{region 'Documentation'}
(*!
<summary>Check that IN is strictly later than Minimum.</summary>
*)
{endregion}
FUNCTION_BLOCK AssertLaterThan_Time EXTENDS AssertionBase
VAR_INPUT
    IN : TIME; //! Actual value checked or observed by this Assertion.
    Minimum : TIME; //! Exclusive lower bound; the actual value or count must be greater.
END_VAR

SUPER^();

{region 'Documentation'}
(*!
<summary>Evaluate the typed duration relation and report higher-priority errors first.</summary>
*)
{endregion}
METHOD PROTECTED Assert
VAR
    Message : STRING(GVL_Constants.MessageLength);
    MinimumText : STRING(GVL_Constants.AssertionValueLength);
    ActualText : STRING(GVL_Constants.AssertionValueLength);
END_VAR
IF NOT EvaluationActive THEN
    RETURN;
END_IF;

IF Result = E_Result.Error THEN
    RETURN;
END_IF;

IF Result = E_Result.Failed THEN
    RETURN;
END_IF;

IF IN <= Minimum THEN
    MinimumText := TIME_TO_STRING(Minimum);
    ActualText := TIME_TO_STRING(IN);
    Message := CONCAT('Assertion failed: value is not later than limit. Minimum = ',
        MinimumText);
    Message := CONCAT(Message, ', Actual = ');
    Message := CONCAT(Message, ActualText);
    Message := CONCAT(Message, '.');
    Fail(Message := Message);
    RETURN;
END_IF;

Pass();
END_METHOD

END_FUNCTION_BLOCK

(* stored: Version 1.1.0.1
   POU AssertLaterThan_Time: Id {9ff3d36c-af1e-41ef-b888-d1db9372648d}, SpecialFunc None
   Folder Internal: Id {66555888-7264-4976-86bf-22a5f2c839ba}
   Method Assert: Id {b7093085-d7a7-4d33-890b-31927c488bc4} *)
